(* PLC project TankControl, plcforge plcforge examples 0.4.0 *)
(* stored: creationDateTime 2026-02-18T11:40:00 *)

(* Level control for a buffer tank with an overfill alarm. *)
FUNCTION_BLOCK TankControl
  VAR_INPUT
    level : REAL;  (* Measured level in percent *)
    lowSetpoint : REAL := 20.0;  (* Pump starts below this level *)
    highSetpoint : REAL := 80.0;  (* Pump stops above this level *)
  END_VAR
  VAR_OUTPUT
    pump : BOOL;  (* Feed pump contactor *)
    overfillAlarm : BOOL;  (* Level stayed above the high setpoint for too long *)
  END_VAR
  VAR
    pumpLatch : RS;
    overfillTimer : TON;
  END_VAR
  VAR  (* added by the conversion: wires and edge detectors of the diagram *)
    _LT4_OUT : BOOL;
    _GT5_OUT : BOOL;
  END_VAR

(* FBD diagram, written out as Structured Text *)
pumpLatch(S := _LT4_OUT, R1 := _GT5_OUT);
pump := pumpLatch.Q1;
overfillTimer(IN := _GT5_OUT, PT := T#3s);
overfillAlarm := overfillTimer.Q;
_LT4_OUT := level < lowSetpoint;
_GT5_OUT := level > highSetpoint;
END_FUNCTION_BLOCK
